(*
SPDX-FileCopyrightText: c 2026 Oleksandr Tiutyk <trofimich@gmail.com>
SPDX-License-Identifier: MIT
License: https://opensource.org/license/mit
*)

(*!
<summary>Checks live changes of referenced engineering and raw limits.</summary>
<description>
Uses fresh method-local fixtures in a single task cycle.
</description>
*)

{attribute 'no_assign'}
{attribute 'no_explicit_call' := 'do not call this function block directly'}
FUNCTION_BLOCK DynamicRangeAnalogValueConverterTest EXTENDS TOF_Testing.SingleCycleTest
VAR_STAT
	{attribute 'hide'}
	_ClassName : STRING := __POUNAME();
END_VAR

(*!
<summary>Checks live changes of referenced engineering and raw limits.</summary>
*)
METHOD PROTECTED ExecuteTest
VAR
	minimumEngineeringValue : LREAL := 0.0;
	maximumEngineeringValue : LREAL := 100.0;
	minimumRawValue : TOF_Devices_IO.RAW_ANALOG_VALUE;
	maximumRawValue : TOF_Devices_IO.RAW_ANALOG_VALUE;
	converter : TOF_Devices_IO.DynamicRangeAnalogValueConverter(
		minAnalogValue := minimumEngineeringValue,
		maxAnalogValue := maximumEngineeringValue,
		minRawValue := minimumRawValue,
		maxRawValue := maximumRawValue
	);
	rawResult : TOF_Devices_IO.RAW_ANALOG_VALUE;
END_VAR
minimumRawValue.Int32 := 0;
minimumRawValue.Int16 := 0;
maximumRawValue.Int32 := 0;
maximumRawValue.Int16 := 1000;

rawResult := converter.ConvertAnalogValueToRawValue(
	analogValue := 50.0,
	rawValueType := TOF_Devices_IO.RAW_ANALOG_VALUE_TYPE.INT16
);
Assert.ThatInt(
	actual := rawResult.Int16,
	message := "Initial dynamic scale"
).ToBe(expected := 500);

// Change the referenced engineering limit.
maximumEngineeringValue := 200.0;

rawResult := converter.ConvertAnalogValueToRawValue(
	analogValue := 50.0,
	rawValueType := TOF_Devices_IO.RAW_ANALOG_VALUE_TYPE.INT16
);
Assert.ThatInt(
	actual := rawResult.Int16,
	message := "Dynamically updated scale"
).ToBe(expected := 250);

maximumRawValue.Int16 := INT#2000;
rawResult := converter.ConvertAnalogValueToRawValue(
	analogValue := LREAL#50.0,
	rawValueType := TOF_Devices_IO.RAW_ANALOG_VALUE_TYPE.INT16
);

Assert.ThatInt(
	actual := rawResult.Int16,
	message := "Changing the referenced raw maximum must update the scale"
).ToBe(expected := INT#500);
END_METHOD

//! <summary>Borrows the concrete class name. Callers must not modify it.</summary>
{attribute 'monitoring' := 'call'}
PROPERTY ClassName : REFERENCE TO STRING
GET
ClassName REF= _ClassName;
END_GET
END_PROPERTY

//! <summary>Borrows the compiler-initialized namespace name. Callers must not modify it.</summary>
{attribute 'monitoring' := 'call'}
PROPERTY NamespaceName : REFERENCE TO STRING
GET
NamespaceName REF= CurrentNamespace.Name;
END_GET
END_PROPERTY

//! <summary>Reports the concrete instance size in bytes.</summary>
{attribute 'monitoring' := 'call'}
PROPERTY SelfSize : ULINT
GET
SelfSize := XSIZEOF(THIS^);
END_GET
END_PROPERTY

END_FUNCTION_BLOCK

(* stored: Version 1.1.0.1
   POU DynamicRangeAnalogValueConverterTest: Id {0f28cc33-5f83-4818-9a0c-a90b49419956}, SpecialFunc None
   Method ExecuteTest: Id {450ccd1e-e6a9-4ba8-93a3-a1cad96bbdf9}
   Property ClassName: Id {f3111f2f-bff8-4fa1-8680-735bfe65aeba}
   Get Get: Id {2a3e0426-407e-44e1-b9ad-1541f793b400}
   Property NamespaceName: Id {3f2e59d1-1dc9-4c20-9461-bdda43db5862}
   Get Get: Id {0ff83154-0e50-4841-bb11-d32dfebbeaea}
   Property SelfSize: Id {900bec67-b843-4846-a959-facd350d2a13}
   Get Get: Id {32965159-cbdf-4aab-99ef-00f10b2dc30f} *)
